(* CODESYS project twincat-tools.library
   Author: hganchev
   Placeholder: tc-tools
   Title: tc-tools
   Version: 1.0.0.0
   DefaultNamespace: tc-tools
   Company: hganchev

Project tree, tasks and I/O mapping:
  libraries: Tc2_Standard, * (Beckhoff Automation GmbH); Tc2_System, * (Beckhoff Automation GmbH); Tc2_Utilities, * (Beckhoff Automation GmbH); Tc3_Module, * (Beckhoff Automation GmbH); TcUnit, * (www.tcunit.org)
  DUTs/
  Examples/
    ExportREALData/
      function block ExportRealDataToFile [ST]
  GVLs/
    global variables Parameters
  POUs/
    Export/
      function block ExportArrayREALDataToTextFile [ST]
    Round/
      function F_ROUNDLREAL [ST]
      function F_ROUNDREAL [ST]
    String/
      function F_STRINGSPLIT [ST]
    TimeStamp/
      function F_GETTIMESTAMP [ST]
  Version/
    global variables Global_Version
  VISUs/
*)

// GVLs/Parameters
{attribute 'qualified_only'}
VAR_GLOBAL CONSTANT
	sNewLineSymbol			: STRING(3) := '$0A'; 	// Control character new line, corresponds to '$L' and '$SN'
	sLineBreakSymbol		: STRING(3) := '$0D';	// Control character line break, corresponds to '$R'
	
	// Export Array REAL data to text file parameters
	iArrayREALSize						: INT := 255;
	diByteMultiplierForExport			: DINT := 10; // This multiplies with array Size
	
	// Split Parameters
	iSplitArraySize						: INT := 4;
END_VAR

// Version/Global_Version
{attribute 'TcGenerated'}
{attribute 'no-analysis'}
{attribute 'linkalways'}
// This function has been automatically generated from the project information.
VAR_GLOBAL CONSTANT
	{attribute 'const_non_replaced'}
	stLibVersion_tc_tools : ST_LibVersion := (iMajor := 1, iMinor := 0, iBuild := 0, iRevision := 0, nFlags := 0, sVersion := '1.0.0.0');
END_VAR

// Examples/ExportREALData/ExportRealDataToFile
FUNCTION_BLOCK ExportRealDataToFile
VAR_INPUT
	arrREALData				: ARRAY[0..Parameters.iArrayREALSize] OF REAL;
	sFilePath				: STRING(255); // File Path
	bUseTimeStamp 			: BOOL;
	bRoundREALDataValues	: BOOL;
	iRoundingDecIndex		: INT := 2; 
	
	bExport					: BOOL;
END_VAR
VAR_OUTPUT
	bExportDone					: BOOL; // Trigger signal for ExportDone
END_VAR
VAR	
	sInputFilePath			: STRING(255);
	// TimeStamp
	timeStamp				: STRING(255);
	sFilePathPlusTimestamp	: STRING(255);
	fbSysTime   			: FB_LocalSystemTime := ( bEnable := TRUE, dwCycle := 1 );
	
	// Export Data
	fbExport 				: ExportArrayREALDataToTextFile;
	
	i						: INT;
END_VAR

// get system time
fbSysTime();

// use time stamp to file name
IF bUseTimeStamp THEN
	// get time stamp
	timeStamp := F_GETTIMESTAMP(fbSysTime.systemTime, '_', '_');
	sFilePathPlusTimestamp := INSERT(sFilePath,CONCAT('_',timeStamp),FIND(sFilePath, '.txt') - 1);
	sInputFilePath := sFilePathPlusTimestamp;
ELSE
	sInputFilePath := sFilePath;
END_IF

// round array data values
IF bRoundREALDataValues THEN
	FOR i := 0 TO Parameters.iArrayREALSize DO
		arrREALData[i] := F_ROUNDREAL(arrREALData[i], iRoundingDecIndex);
	END_FOR
END_IF


fbExport(
	arrData:= arrREALData, 
	bExecute:= bExport, 
	bUseTimeStamp:= bUseTimeStamp, 
	sFilePath:= sInputFilePath, 
	bDone=> bExportDone);

END_FUNCTION_BLOCK

// POUs/TimeStamp/F_GETTIMESTAMP
FUNCTION F_GETTIMESTAMP : STRING(255)
VAR_INPUT
	systemTime				: TIMESTRUCT;			// Using Tc2_Utilities to have the TIMESTRUCT
	strSeparatorDate		: STRING(1) := '_';		// Separator between Year,Month,Day
	strSeparatorTime		: STRING(1) := ':';		// Separator between Hours, Minutes, Seconds		
END_VAR
VAR
	stYear					: STRING;
	stMonth					: STRING;
	stDay					: STRING;
	stHours					: STRING;
	stMinutes				: STRING;
	stSeconds				: STRING;
END_VAR

stYear 		:= CONCAT(WORD_TO_STRING(systemTime.wYear), strSeparatorDate);
stMonth		:= CONCAT(WORD_TO_STRING(systemTime.wMonth), strSeparatorDate);
stDay 		:= CONCAT(WORD_TO_STRING(systemTime.wDay), strSeparatorDate);
stHours 	:= CONCAT(WORD_TO_STRING(systemTime.wHour), strSeparatorTime);
stMinutes 	:= CONCAT(WORD_TO_STRING(systemTime.wMinute), strSeparatorTime);
stSeconds 	:= WORD_TO_STRING(systemTime.wSecond);
F_GETTIMESTAMP := CONCAT(stYear,CONCAT(stMonth,CONCAT(stDay,CONCAT(stHours,CONCAT(stMinutes,stSeconds)))));

END_FUNCTION

// POUs/Round/F_ROUNDREAL
FUNCTION F_ROUNDREAL : REAL
VAR_INPUT
	rValue		: REAL; // Input Value
	iDecNumber	: INT; 	// Numbers after decimal point
END_VAR
VAR
	rOutValue	: REAL;
	rLeftValue	: REAL;
END_VAR

rOutValue := rValue * EXPT(10,iDecNumber);
rLeftValue := rOutValue - TRUNC(rOutValue);
IF rLeftValue >= 0.5 THEN
	rOutValue := TRUNC(rOutValue + 1) / EXPT(10,iDecNumber);
ELSE
	rOutValue := TRUNC(rOutValue) / EXPT(10,iDecNumber);
END_IF
F_ROUNDREAL := rOutValue;

END_FUNCTION

// POUs/Export/ExportArrayREALDataToTextFile
FUNCTION_BLOCK ExportArrayREALDataToTextFile
VAR_INPUT
	arrData 				: ARRAY[0..Parameters.iArrayREALSize] OF REAL;
	bExecute				: BOOL;
	bUseTimeStamp			: BOOL;
	sFilePath				: STRING(255) := 'C:\data.txt';
END_VAR         			
VAR_OUTPUT      			
	bDone					: BOOL;
END_VAR
VAR
	fileOpen				: FB_FileOpen;
//	fileWrite				: FB_FilePuts;
	fileWrite				: FB_FileWrite;
	fileClose				: FB_FileClose;
	                		
	fileHandle				: UINT;
	nSizeWritten			: UDINT;
	
	arrayDataByte			: ARRAY[0..iArrayByteSize] OF BYTE;
	sData					: ARRAY[0..Parameters.iArrayREALSize] OF STRING(255);

	i						: INT;
	j						: INT;
	k						: DINT;	// track of byte array
END_VAR

VAR CONSTANT
	iArrayByteSize 			: DINT := Parameters.diByteMultiplierForExport * Parameters.iArrayREALSize;
END_VAR

bDone := FALSE;
fileClose(bExecute := FALSE);

// file write init
fileWrite(tTimeout:= T#2S);

IF bExecute	THEN	
	// open file
	fileOpen(sPathName := sFilePath, nMode := FOPEN_MODEWRITE,
		 ePath := PATH_GENERIC, hFile => fileHandle, bExecute := TRUE);
		 
	// Clear data
	MEMSET(ADR(arrayDataByte), 16#00, SIZEOF(arrayDataByte));
	
	k := 0;
	// Prepare string data 
	FOR i := 0 TO Parameters.iArrayREALSize DO
		sData[i] := REAL_TO_STRING(arrData[i]);
		IF i > 0 THEN
			sData[i] := CONCAT(Parameters.sNewLineSymbol,sData[i]);
		END_IF
		// Convert to byte for every sData symbol
		FOR j := 0 TO LEN(sData[i]) DO
			MEMCPY(ADR(arrayDataByte[k]),ADR(sData[i][j]), 1);
			k := k + 1;
		END_FOR
	END_FOR
	
	// Write Data
	IF fileHandle <> 0 THEN
		fileWrite(	hFile:= fileHandle, 
					pWriteBuff:= ADR(arrayDataByte), 
					cbWriteLen:= SIZEOF(arrayDataByte), 
					bExecute := TRUE);
	END_IF
	
	IF fileWrite.cbWrite > 0 THEN
		bDone := TRUE;
	END_IF
ELSIF NOT bExecute THEN
	IF NOT fileWrite.bBusy THEN
		fileWrite(bExecute := FALSE);
		fileOpen(bExecute := FALSE);
		fileClose(hFile := fileHandle, bExecute := TRUE);
	END_IF
END_IF

END_FUNCTION_BLOCK

// POUs/Round/F_ROUNDLREAL
FUNCTION F_ROUNDLREAL : LREAL
VAR_INPUT
	rValue		: LREAL; // Input Value
	iDecNumber	: INT; 	// Numbers after decimal point
END_VAR
VAR
	rOutValue	: LREAL;
	rLeftValue	: LREAL;
END_VAR

rOutValue := rValue * EXPT(10,iDecNumber);
rLeftValue := rOutValue - TRUNC(rOutValue);
IF rLeftValue >= 0.5 THEN
	rOutValue := TRUNC(rOutValue + 1) / EXPT(10,iDecNumber);
ELSE
	rOutValue := TRUNC(rOutValue) / EXPT(10,iDecNumber);
END_IF
F_ROUNDLREAL := rOutValue;

END_FUNCTION

// POUs/String/F_STRINGSPLIT
FUNCTION F_STRINGSPLIT : ARRAY[0..Parameters.iSplitArraySize] OF STRING(255)
VAR_INPUT
	sInput			: STRING(255);
	sSplitChar		: STRING(1);
END_VAR
VAR
	sCopy			: STRING(255);
	sSplit			: STRING(255);
	iDeleteLen		: INT;
	i				: INT;
END_VAR

sCopy := sInput;

FOR i := 0 TO Parameters.iSplitArraySize DO
	IF FIND(sCopy, sSplitChar) > 0 THEN
		sSplit := LEFT(sCopy, FIND(sCopy, sSplitChar) - 1);
		iDeleteLen := LEN(sSplit) + LEN(sSplitChar);
	ELSE
		sSplit := sCopy;
		iDeleteLen := LEN(sSplit);
	END_IF
	
	// Take the string value
	F_STRINGSPLIT[i] := sSplit;
	
	// Delete 
	sCopy := DELETE(sCopy, iDeleteLen, 1);
	
	// End of split
	IF sCopy = '' THEN
		EXIT;
	END_IF
END_FOR

END_FUNCTION
